Staubli VAL3: waitDigInput.pgx

public program waitDigInput(dio x_dIn, bool x_bValue, bool& x_bError)
  local string l_sDesc
  local string l_sPath
begin
  if ioStatus(x_dIn,l_sDesc,l_sPath)>=0
    x_bError=false
    wait(x_dIn==x_bValue)
  else
    x_bError=true
    logMsg("通信终端，等待通信恢复")
    wait(x_dIn==x_bValue)
    logMsg("通信已恢复")
    //    logMsg("Signal "+l_sPath+" error."+"Description:"+l_sDesc)
  endIf
end
